Fanuc KAREL source: KA00210.KL

PROGRAM KA00210
%NOLOCKGROUP
VAR
  SRC: ARRAY[4] OF XYZWPR
  DST: ARRAY[4] OF BOOLEAN
BEGIN
  DST = SRC
END KA00210
